Staubli VAL3: iolink.pgx

public program iolink()
  local num l_i
begin
  for l_i = 0 to size(O_safePoint)-1
    dioLink(O_safePoint[l_i],io:dOutput[nIO_spindex[l_i]])
  endFor

  for l_i =0 to size(O_safeZone)-1
    dioLink(O_safeZone[l_i],io:dOutput[nIO_Zoneindex[l_i]])
  endFor
end
